(* IEC 61131-3 sources: rusty/compiler/plc_cfc/fixtures/execution_control/valid/enable_from_function, 2 files *)

(* ---- isNonZero.st ---- *)
FUNCTION isNonZero : BOOL
VAR_INPUT
    val : DINT;
END_VAR
    isNonZero := val <> 0;
END_FUNCTION

(* ---- safeDiv.st ---- *)
FUNCTION safeDiv : DINT
VAR_INPUT
    dividend : DINT;
    divisor : DINT;
END_VAR
    safeDiv := dividend / divisor;
END_FUNCTION
